Fanuc KAREL source: KT00819.KL

PROGRAM KT00819
%NOLOCKGROUP
VAR
  S1: STRING[80]
  S2: STRING[80]
  OUT: REAL
BEGIN
  S1 = 'A'
  S2 = 'B'
  S1 = 'A'
  S2 = 'B'
  OUT = LN(S1)
END KT00819
